Staubli VAL3: init.pgx

public program init()
begin
  //更改_nPuleStartClk的大小
  if size(_nPuleStartClk)!=io:nMaxdigital
    resize(_nPuleStartClk,1,io:nMaxdigital)
    libSave()
  endIf
  //num
  _nActStackIndex=0
  //Bool
  bPushToStack=false
  //
  call clearActStack()
  //
  setMoveId(0)
end
